SUBAPPLICATION Uebung_094b5_AX (* Wie Uebung_094b_AX, aber mit AOption_AD_DEMUX_2 (Bitmaske, Multi-Select) statt AOption_AUI_DEMUX_2 (Index, Single-Select): Bit0 schaltet OptionalGroup_001, Bit1 schaltet OptionalGroup_002 - beide koennen hier gleichzeitig aktiv sein. *)
  (* Standard: 61499-2; Description: Copyright (c) 2026 Meisterschulen am Ostbahnhof This program and the accompanying materials are made available under the terms of the Eclipse Public License 2.0 which is available at https://www.eclipse.org/legal/epl-2.0/ SPDX-License-Identifier: EPL-2.0 *)
  (* Version 1.0, 2026-10-13, Franz Höpfinger, Meisterschulen am Ostbahnhof, Kopie von Uebung_094b_AX, AD_TO_AUI+AUI_TO_AUI2 durch AD_TO_AD2 ersetzt (kein Zwischenschritt noetig, da NumericValue_IDA.IN bereits DWORD/AD ist) und AOption_AUI_DEMUX_2 durch AOption_AD_DEMUX_2 ersetzt. *)
  PACKAGE Uebungen;
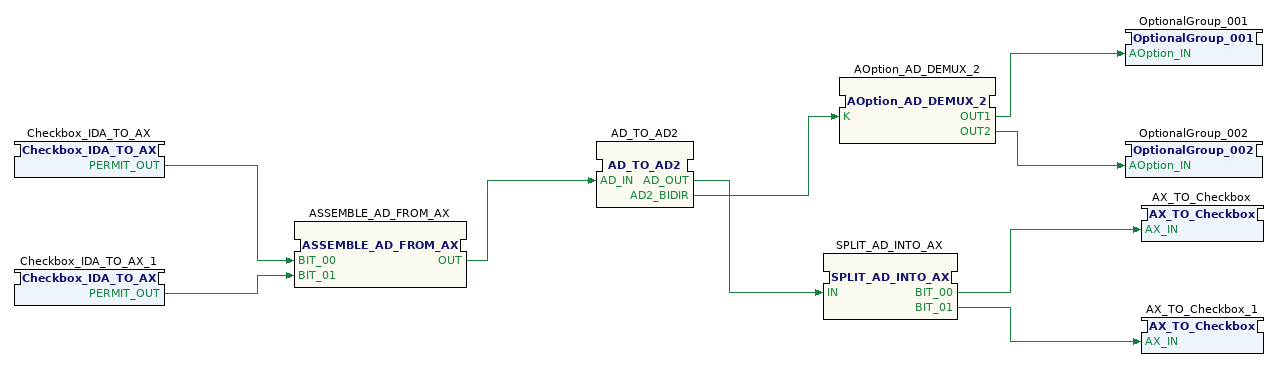
  FBS
    AOption_AD_DEMUX_2 : Option::selection::AOption_AD_DEMUX_2;
    AD_TO_AD2 : adapter::conversion::bidirectional::AD_TO_AD2;
    SPLIT_AD_INTO_AX : adapter::splitting::SPLIT_AD_INTO_AX;
    ASSEMBLE_AD_FROM_AX : adapter::assembling::ASSEMBLE_AD_FROM_AX;
  END_FBS
  SUBAPPS
    OptionalGroup_001 : MyLib_AX_Option::sys::OptionalGroup_001;
    OptionalGroup_002 : MyLib_AX_Option::sys::OptionalGroup_002;
    Checkbox_IDA_TO_AX : MyLib::sys::Checkbox_IDA_TO_AX;
    Checkbox_IDA_TO_AX_1 : MyLib::sys::Checkbox_IDA_TO_AX;
    AX_TO_Checkbox : MyLib::sys::AX_TO_Checkbox;
    AX_TO_Checkbox_1 : MyLib::sys::AX_TO_Checkbox;
  END_SUBAPPS
  ADAPTER_CONNECTIONS
    AOption_AD_DEMUX_2.OUT1 TO OptionalGroup_001.AOption_IN;
    AOption_AD_DEMUX_2.OUT2 TO OptionalGroup_002.AOption_IN;
    ASSEMBLE_AD_FROM_AX.OUT TO AD_TO_AD2.AD_IN;
    AD_TO_AD2.AD_OUT TO SPLIT_AD_INTO_AX.IN;
    AD_TO_AD2.AD2_BIDIR TO AOption_AD_DEMUX_2.K;
    Checkbox_IDA_TO_AX.PERMIT_OUT TO ASSEMBLE_AD_FROM_AX.BIT_00;
    Checkbox_IDA_TO_AX_1.PERMIT_OUT TO ASSEMBLE_AD_FROM_AX.BIT_01;
    SPLIT_AD_INTO_AX.BIT_00 TO AX_TO_Checkbox.AX_IN;
    SPLIT_AD_INTO_AX.BIT_01 TO AX_TO_Checkbox_1.AX_IN;
  END_CONNECTIONS
END_SUBAPPLICATION
